// Settable I_SafetyDiagnostics for tests of consumers (HMI gateway): the properties return the inputs.
FUNCTION_BLOCK FB_SafetyDiagnosticsStub IMPLEMENTS BROTLib.I_SafetyDiagnostics
VAR_INPUT
	bStoActive		: BOOL;
	bRestartPending	: BOOL;
	stItems			: BROTLib.ST_SafetyItems;
END_VAR

PROPERTY StoActive : BOOL
GET
StoActive := bStoActive;
END_GET
END_PROPERTY

PROPERTY RestartPending : BOOL
GET
RestartPending := bRestartPending;
END_GET
END_PROPERTY

PROPERTY Items : BROTLib.ST_SafetyItems
GET
Items := stItems;
END_GET
END_PROPERTY

END_FUNCTION_BLOCK

(* stored: Version 1.1.0.1, ProductVersion 3.1.4024.15
   POU FB_SafetyDiagnosticsStub: Id {5b52800c-fc81-42ef-9d5a-d5ab5f2cee2b}, SpecialFunc None
   Property StoActive: Id {cd3f9f17-d496-4716-b47d-0268b7faf947}
   Get Get: Id {f438f7bd-6b50-4f06-ace2-b20fea1df5a6}
   Property RestartPending: Id {9ae9f196-9513-418e-94a1-049297f5ae9e}
   Get Get: Id {c17a25c5-9e18-42f8-89d4-37290332a1eb}
   Property Items: Id {67236ac8-e6e2-4a7f-a8b9-eb7013295204}
   Get Get: Id {ac8256a4-9b63-449a-ac0e-7862a9a05128} *)
